// Exact current capability identity/type/revision; no blanket stale migration.
// AnyRevision: a restored document carries the ConfigRev of an earlier run, which
// says nothing about this one; the per-record identity, type and revision still do.
METHOD PRIVATE _M_ValidateSetShape : BOOL
VAR_INPUT
    Store : I_ConfigStore;
    Info : ST_ConfigSetInfo;
    AnyRevision : BOOL;
END_VAR
VAR
    expectedInfo : ST_ConfigSetInfo;
    expected : ST_ConfigRecord;
    record : ST_ConfigRecord;
    i : INT;
    j : INT;
    hits : INT;
END_VAR
_M_ValidateSetShape := FALSE;
IF (Store = 0) OR (Info.RootIdentity <> Status.Name)
OR (Info.SetSchema <> CONFIG_SET_SCHEMA)
OR (Info.RecordCount < 1) OR (Info.RecordCount > PL_Fraktal.MAX_SET_RECORDS) THEN
    _M_RejectConfigSet(Scope := Info.RootIdentity, Key := Info.SetName); RETURN;
END_IF
IF NOT AnyRevision AND ((Info.ConfigRev = 0) OR (Info.ConfigRev > ConfigRev)) THEN
    _M_RejectConfigSet(Scope := Info.RootIdentity, Key := Info.SetName); RETURN;
END_IF
IF NOT _snapshot.M_ReadInfo(SetName := '_validation', Info := expectedInfo) THEN RETURN; END_IF

FOR i := 1 TO Info.RecordCount DO
    IF NOT Store.M_ReadRecord(SetName := Info.SetName, Index := i, Record := record) THEN RETURN; END_IF
    hits := 0;
    FOR j := 1 TO expectedInfo.RecordCount DO
        _snapshot.M_ReadRecord(SetName := '_validation', Index := j, Record := expected);
        IF (record.Scope = expected.Scope) AND (record.WriteKey = expected.WriteKey) THEN
            IF (record.Kind <> expected.Kind) OR (record.ValueType <> expected.ValueType)
            OR (record.Revision <> expected.Revision) THEN
                _M_RejectConfigSet(Scope := record.Scope, Key := record.WriteKey); RETURN;
            END_IF
            hits := hits + 1;
        END_IF
    END_FOR
    IF hits <> 1 THEN
        _M_RejectConfigSet(Scope := record.Scope, Key := record.WriteKey); RETURN;
    END_IF
END_FOR
// Station sets may carry a subset; a Model bank or Line calendar is complete.
IF (Info.Kind <> E_ConfigKind.STATION_CFG) AND (Info.RecordCount <> expectedInfo.RecordCount) THEN
    _M_RejectConfigSet(Scope := Info.RootIdentity, Key := Info.SetName); RETURN;
END_IF
_M_ValidateSetShape := TRUE;
END_METHOD

// Append an inactive provider record. Live recipe and existing ordinals stay fixed.
METHOD CreateModel : BOOL
VAR_INPUT
    ModelCode : STRING(160);
    SourceIndex : UDINT;
    FromSet : BOOL;
    SetName : STRING(80);
END_VAR
VAR
    i : INT;
    info : ST_ConfigSetInfo;
    record : ST_ConfigRecord;
    source : I_ConfigStore;
    sourceName : STRING(80);
END_VAR
CreateModel := FALSE;
IF NOT _M_ConfigRestored() THEN
    RETURN;
END_IF
_exportNext := 0;
_M_SyncModelCatalog();
IF (_modelCatalog = 0) OR (_pModelRegion = 0) OR (_modelRegionSize < SIZEOF(UINT))
OR (ModelCode = '') OR (LEN(ModelCode) > 64) OR (AvailableModelCount >= ModelCapacity)
OR NOT Access.PermitsLogged(Gate := E_GatedAction.CONFIG_SET) THEN RETURN; END_IF
FOR i := 1 TO AvailableModelCount DO
    IF AvailableModels[i].ModelCode = ModelCode THEN RETURN; END_IF
END_FOR
// The exact bytes being validated are copied into the existing view buffer.
IF NOT _M_CaptureConfig(SetName := '_validation', Kind := E_ConfigKind.PAR_CFG,
        ModelIndex := SourceIndex) THEN RETURN; END_IF
source := _snapshot;
sourceName := '_validation';
IF FromSet THEN
    IF _configStore = 0 THEN RETURN; END_IF
    IF NOT _M_CopySet(SetName := SetName) THEN RETURN; END_IF
    IF NOT _loadSnapshot.M_ReadInfo(SetName := SetName, Info := info) THEN RETURN; END_IF
    IF info.Kind <> E_ConfigKind.PAR_CFG THEN RETURN; END_IF
    IF NOT _M_ValidateSetShape(Store := _loadSnapshot, Info := info,
            AnyRevision := FALSE) THEN RETURN; END_IF
    source := _loadSnapshot;
    sourceName := SetName;
END_IF
IF NOT source.M_ReadInfo(SetName := sourceName, Info := info) THEN RETURN; END_IF
MEMCPY(destAddr := ADR(_modelBuf), srcAddr := _pModelRegion, n := _modelRegionSize);
IF SourceIndex > 0 THEN
    IF AvailableModels[SourceIndex].ModelCode <> Model.ModelCode THEN
    IF NOT _modelProvider.Load(ModelCode := AvailableModels[SourceIndex].ModelCode,
            RecipeKey := _modelKey, pParCfg := ADR(_modelBuf), Size := _modelRegionSize) THEN RETURN; END_IF
    END_IF
END_IF
_pModelView := ADR(_modelBuf);
FOR i := 1 TO info.RecordCount DO
    IF NOT source.M_ReadRecord(SetName := sourceName, Index := i, Record := record) THEN EXIT; END_IF
    // A provider with one root record cannot clone another owner's recipe bank.
    IF NOT _M_OwnsModelRecord(Record := record) THEN EXIT; END_IF
    IF NOT Access.M_PermitsLevelLogged(Required := _M_DataLevelOf(TargetPath := record.Scope,
            WriteKey := record.WriteKey, ForWrite := FALSE)) THEN EXIT; END_IF
    IF NOT Access.M_PermitsLevelLogged(Required := _M_DataLevelOf(TargetPath := record.Scope,
            WriteKey := record.WriteKey, ForWrite := TRUE)) THEN EXIT; END_IF
    IF NOT SUPER^.M_ApplyConfigWrite(Scope := record.Scope, WriteKey := record.WriteKey,
            Revision := record.Revision, TextValue := record.ValueText, RootReady := TRUE) THEN EXIT; END_IF
END_FOR
_pModelView := 0;
IF i <= info.RecordCount THEN RETURN; END_IF
CreateModel := _modelCatalog.M_CreateModel(ModelCode := ModelCode, RecipeKey := _modelKey,
    pData := ADR(_modelBuf), Size := _modelRegionSize);
IF CreateModel THEN
    _M_SyncModelCatalog();
    _M_MarkPersistPending();
END_IF
END_METHOD

METHOD ExportCurrentConfig : BOOL
VAR_INPUT
    SetName : STRING(80);
    Kind : E_ConfigKind;
    ModelIndex : UDINT;
    Token : STRING(160);
END_VAR
VAR
    info : ST_ConfigSetInfo;
    record : ST_ConfigRecord;
    i : INT;
END_VAR
ExportCurrentConfig := FALSE;
_exportNext := 0;
ConfigSetDocument := '';
ConfigSetDocumentLines := 0;
IF (Token = '') OR Access.ReqLogout
OR NOT Access.Permits(Gate := E_GatedAction.CONFIG_SET) THEN RETURN; END_IF
IF NOT _M_CaptureConfig(SetName := SetName, Kind := Kind, ModelIndex := ModelIndex) THEN RETURN; END_IF
_snapshot.M_ReadInfo(SetName := SetName, Info := info);
FOR i := 1 TO info.RecordCount DO
    _snapshot.M_ReadRecord(SetName := SetName, Index := i, Record := record);
    IF NOT Access.M_PermitsLevel(Required := _M_DataLevelOf(TargetPath := record.Scope,
            WriteKey := record.WriteKey, ForWrite := FALSE)) THEN RETURN; END_IF
END_FOR
_exportToken := Token;
_exportSession := Access.SessionGeneration;
_exportName := SetName;
_exportNext := 1;
ConfigSetDocument := _setJson.M_Header(Info := info);
ConfigSetDocumentLine := 0;
ConfigSetDocumentLines := info.RecordCount;
ExportCurrentConfig := ConfigSetDocument <> '';
END_METHOD

METHOD PRIVATE _M_ExportSnapshotLine : BOOL
VAR_INPUT
    SetName : STRING(80);
    Line : INT;
    Token : STRING(160);
END_VAR
VAR
    info : ST_ConfigSetInfo;
    record : ST_ConfigRecord;
END_VAR
_M_ExportSnapshotLine := FALSE;
ConfigSetDocument := '';
ConfigSetDocumentLines := 0;
IF (_exportNext = 0) OR (Line <> _exportNext) OR (Token <> _exportToken)
OR (_exportSession <> Access.SessionGeneration) OR (SetName <> _exportName)
OR Access.ReqLogout
OR NOT Access.Permits(Gate := E_GatedAction.CONFIG_SET) THEN
    _exportNext := 0; RETURN;
END_IF
IF NOT _snapshot.M_ReadInfo(SetName := SetName, Info := info)
OR NOT _snapshot.M_ReadRecord(SetName := SetName, Index := Line, Record := record) THEN
    _exportNext := 0; RETURN;
END_IF
IF NOT Access.M_PermitsLevel(Required := _M_DataLevelOf(TargetPath := record.Scope,
        WriteKey := record.WriteKey, ForWrite := FALSE)) THEN
    _exportNext := 0; RETURN;
END_IF
ConfigSetDocument := _setJson.M_Record(Record := record);
ConfigSetDocumentLine := Line;
ConfigSetDocumentLines := info.RecordCount;
_exportNext := _exportNext + 1;
IF Line = info.RecordCount THEN _exportNext := 0; END_IF
_M_ExportSnapshotLine := ConfigSetDocument <> '';
END_METHOD

END_FUNCTION_BLOCK

(* stored: Version 1.1.0.1, ProductVersion 3.1.4024.16
   POU FB_UnitBase: Id {116d9026-fbad-4cf8-8b52-50d17613c706}, SpecialFunc None
   Method _M_AddReason: Id {63c5e93f-708a-4c3a-aa1b-ee43d815fb4a}
   Method _M_AppendInterlocks: Id {2bc971ff-4cee-49e6-a29f-4f727818205b}
   Method _M_AppendManualInterlocks: Id {c18caeb9-871a-4a4c-aad2-2711e3ced37a}
   Method _M_AppendDecisionInterlocks: Id {bbac41d9-35ba-4800-af52-51cd30b49db7}
   Method _M_AskDecision: Id {4e23ce8a-174c-4663-9cbe-be702ba37032}
   Method _M_ClearDecisionState: Id {db09e3d9-4427-4607-8a90-66b39812e37b}
   Method _M_DecisionCyclic: Id {ff058255-d664-4ce3-986d-8ad7a970388c}
   Method _M_DecisionMatches: Id {2ca48458-620f-4a17-b6d1-b5680778bd4e}
   Method _M_LogDecision: Id {eb357477-2029-4b6d-8688-04dc5df5e04b}
   Method _M_ValidateDecision: Id {1229fbc9-7dc8-4907-b878-f6af733f2c09}
   Method _M_Await: Id {098638cb-fc78-4032-9954-0ceffe6b565c}
   Method _M_CascadeMode: Id {3ac20481-72c5-4cd1-88e5-b9f7eb433162}
   Method _M_ClearPending: Id {cb01b1f4-f591-43f7-a826-970be7300b04}
   Method _M_AuditHmiAccepted: Id {f8865f87-3ae7-472e-b775-3408513a4586}
   Method _M_OwnsModulePath: Id {9b8c6045-f404-4484-937e-b0a8f749d8fd}
   Method _M_EndOfCycle: Id {9824e487-d8d3-4cb9-8c78-a6d2fc09a62d}
   Method _M_HandleHmiRequest: Id {63ae9d50-339f-4904-a8ec-81f853aed962}
   Method _M_HostEvent: Id {76fb49ac-f9ea-4e53-8db6-e7e4e756fd84}
   Method _M_InitModePolicy: Id {df8ba8da-c8fa-411c-85c1-392b353d5cfd}
   Method _M_OeeCompute: Id {2991f1a8-70f1-48a9-aa83-352243818d0a}
   Method _M_OeeUpdate: Id {8a4f011d-5d7a-4935-ad26-8a5fbcf63643}
   Method _M_PartAborted: Id {a55c31e8-06f9-4d10-8c26-4e83b7d5c1f2}
   Method _M_PartEvent: Id {f18c2d47-9b53-4e6a-8c02-3a71d5f0b429}
   Method _M_PartProcessed: Id {e91b5a02-73df-4f16-a8d4-1c30fe8a97d2}
   Method _M_PartReceived: Id {58c0a7d9-14be-4f22-8d6a-9b2ef4c1e370}
   Method _M_PartRecord: Id {7be4f6a3-1d20-4c8e-be55-f2a09318d67c}
   Method _M_PartStarted: Id {02a97d1c-6bb5-4f80-9d34-c58b12f04ae6}
   Method _M_PublishStatus: Id {02d44270-09e8-4bc1-97fd-f43dd3fc44f2}
   Method _M_PushHistory: Id {3f9af757-7ef5-4499-8b8d-04dcd97acc93}
   Method _M_RaiseMaintenance: Id {c92e4b71-6d05-4f88-9e3a-2b17d4c8a054}
   Method _M_RouteConfigWrite: Id {4e524daf-e482-4764-8639-e58c1f363aa3}
   Method _M_WriteBaseConfig: Id {c30f39b4-eae4-421d-a415-c6dc3b402679}
   Method _M_RouteForceChannel: Id {301182d5-8822-451a-950c-49d23daf4640}
   Method _M_RouteManual: Id {9fa4e2c2-3f5f-4681-aed5-559f1df0d2c6}
   Method _M_RecordSequenceStep: Id {bae7334e-b67d-46db-a917-aa05f1522e0f}
   Method _M_ResetSequenceRows: Id {3a7e979a-9c02-4e58-aa36-f0627902f8fb}
   Method _M_SequenceAnnotate: Id {981fa92c-f12b-4972-9483-880edfae72c8}
   Method _M_SequenceAnnotationClear: Id {7256d50d-cf16-4906-8e35-fd394563602f}
   Method _M_SetStep: Id {1066dd3c-baf2-43ea-91d5-309ad4ca7878}
   Method _M_StallWalk: Id {ee453cd4-7027-4207-b43e-f1a12367922c}
   Method _M_StepGate: Id {853d1e75-22c1-46fb-9a92-007882839a98}
   Method _M_Supports: Id {5285aa9e-3e18-4090-bed9-0119293228bb}
   Method _M_SupportsRunStyle: Id {f4e81ed4-d8b0-494c-bd7a-6b417d6219cf}
   Method _M_TakeDecision: Id {e2e1443d-0421-4608-8ae5-b7bb44177b3c}
   Method CountGood: Id {852e951b-039f-45bd-80a3-6417310e2406}
   Method CountNok: Id {a686f5b6-4c90-4e12-9d98-fa111d14dfe8}
   Method CountRework: Id {5c8e02d7-9a41-4f36-8b52-e04a71c6d983}
   Method M_AppendConfig: Id {29c7f5d4-0b81-4ae3-9762-84f6d013ba58}
   Method SetConfigStore: Id {1f6b90d4-38a2-4c57-9e01-b47d2c85a3f6}
   Method SetPersistMedium: Id {90949ce0-2dde-4312-82c9-779c3854619d}
   Method SetConfigPersistence: Id {a5c37e08-9412-4bd6-83f9-6e05b17c94a2}
   Method SetConfigPersistWindow: Id {5db2740a-9e18-4c63-b0f5-8a2914e7c036}
   Method SetConfigRestorePolicy: Id {72e4a1b9-c530-46df-8127-93b605ea4d78}
   Method _M_MarkPersistPending: Id {6d09fb35-2a84-41ce-b7f0-58d2e1937a4b}
   Method _M_ConfigPersistFailed: Id {3a81c6e7-40b2-4d95-916f-c82705bd4e13}
   Method _M_ConfigPersistCyclic: Id {9c0d4318-b7a5-42e6-8f13-05ea7c9b2d40}
   Method _M_ConfigRestored: Id {c723ef57-9111-489a-87e1-2e9e98d880fe}
   Method _M_LiveCyclic: Id {aad84a07-4f6e-415a-a949-44d11c57baf2}
   Method _M_LiveReadFailed: Id {c1b391b8-49e2-405b-9490-706629300cca}
   Method _M_LivePassFailed: Id {3fff4db1-40c0-4916-a009-f750b7b16137}
   Method _M_LiveItemUsed: Id {2d7178d4-917d-4032-9b90-b6d8a8215873}
   Method _M_LiveKey: Id {77a63a7d-cd03-4447-be78-e758d5ef1591}
   Method _M_LiveModelsKept: Id {166da471-060a-4724-bca3-30a7b039d62b}
   Method _M_LiveRestoreItem: Id {b20141f1-cfd8-47d0-b996-33c491a3a370}
   Method _M_LiveApply: Id {031ae06a-8d84-4843-bce8-ed6d53fdc0d1}
   Method _M_ModelIndexOf: Id {055b30d9-edd2-408c-ae7f-7015e649658e}
   Method _M_DrainRestoreLoss: Id {0b7e5294-16ad-43c1-a8f6-249d038be715}
   Method _M_AnnounceRestoreLoss: Id {77125c95-ab46-4aaa-9f22-3a07f8e7fd8f}
   Method AcknowledgeConfigRestore: Id {e18c47b3-5029-4ed6-9a71-b3406fc25d89}
   Method _M_RejectConfigSet: Id {5f2a90c6-8b41-4d73-bec0-172e845f39ab}
   Method _M_SetOpAllowed: Id {3d70b95e-c284-41f0-86ba-9e15c703da42}
   Method DeleteConfigSet: Id {e533f05f-2594-42e8-8c99-81d549fc4090}
   Method _M_DataLevelOf: Id {181e4912-d325-4208-982a-bde235412443}
   Method M_DeclareDataClass: Id {b9a4a5ae-9fab-42bd-bc82-7e32dffbd2a9}
   Method SetDataClassLevel: Id {047e7f36-274a-4350-8ad6-b77d4f72cc43}
   Method _M_IsLineKey: Id {59358b2d-9028-416d-b8b1-1699a6cd425f}
   Method M_ApplyConfigWrite: Id {09d95f4a-6281-4745-bbd6-78a379c3dcc0}
   Method M_StageConfigWrite: Id {c033d610-c896-4206-a3ad-81018a4dd465}
   Method M_ApplyCapture: Id {e2ff8450-6122-448e-b867-574b3000edfa}
   Method M_ConfigAccessOf: Id {b5882f05-b837-4f44-ba08-a65bdacad4e2}
   Method M_RegisterModelData: Id {9e19e4d6-5131-4b98-84c6-f84c0e107ced}
   Method _M_OpenModelView: Id {93ccf92c-d752-48c8-af0b-7941488b3430}
   Method WriteModelConfig: Id {2a0d9e3e-ba70-4e09-955f-cec98e39642e}
   Method M_AppendModelConfig: Id {0e6d90bf-ad76-4384-ab12-1767af3d1a4f}
   Method _M_SaveModelData: Id {614f64a8-a7bb-415b-89b6-cd5638516728}
   Method SetLine: Id {b3e3c826-6085-43fe-ab9e-5ee8d63ca7f0}
   Method M_ShiftTick: Id {4606cb81-948b-4fb3-a998-828e0341cdfd}
   Method _M_CloseShift: Id {3589014a-a797-47c8-9c22-164193338f8a}
   Method SaveConfigSet: Id {8a4d1e07-63b9-4c25-90fd-e7285a1cb046}
   Method LoadConfigSet: Id {c93f5b28-047e-41da-b6c1-5820ae74f3d9}
   Method _M_ApplySet: Id {f003cd3e-e4eb-4ec5-b15b-c46e595f4b79}
   Method _M_StageOneRecord: Id {b6014e8d-72c3-49a5-80fe-c1738d92406b}
   Method _M_ConfigSetHalfApplied: Id {47db6015-9a2e-4c38-b7f0-d5216e409a83}
   Method ListConfigSets: Id {2e85d740-c6b1-4930-a5df-08417b3ce629}
   Method ExportConfigSetLine: Id {6c1908fe-b432-4a07-95d8-e2603ba7145c}
   Method ImportConfigSetLine: Id {d0a76321-8e54-4bc9-97a2-3f16054eb7d8}
   Method ImportConfigSetPiece: Id {fe4a451b-e9cc-440c-9ade-c56031168c94}
   Method M_SequenceAskDecision: Id {099b4f9d-bc09-44d1-a376-b2e504dbb242}
   Method M_SequenceAwait: Id {c61669f7-ff2f-475c-915e-c23e673ae50d}
   Method M_SequenceClearDecision: Id {f5e88d63-dd7e-45c7-8fcc-149437ebcb66}
   Method M_SequenceComplete: Id {94f85c2c-bf7e-4679-9ad7-df299f9443e9}
   Method M_SequenceCountGood: Id {7ac5d064-bbc3-4e23-a999-5b1106c18501}
   Method M_SequenceEndOfCycle: Id {2465831e-ce6a-49ba-894a-d94a6e5b730d}
   Method M_SequenceFault: Id {6dcf30ea-273a-4919-b53c-93ee346a0722}
   Method M_SequencePartProcessed: Id {f3fe635f-f0ef-4b80-918f-2af11c08a018}
   Method M_SequencePartReceived: Id {9576ad5e-fef2-4d71-bd9f-075e2fbf7f48}
   Method M_SequencePartRecord: Id {272bc8d6-51f1-4e02-a0f6-834fc34cf443}
   Method M_SequencePartStarted: Id {c34399dc-9677-414b-87a7-da41fec81ce1}
   Method M_SequenceRegister: Id {9c12e1e0-2b54-4710-a719-b7dbb939da2c}
   Method _M_BeginSequenceScan: Id {90d173ad-1ac7-44ea-8963-773d827fd02e}
   Method _M_RestartSequences: Id {a7179c76-6bab-4060-a5d3-1d37fa9ff028}
   Method OnAbort: Id {045fbfe7-105f-49b4-bf25-f60661612052}
   Method OnAbortInError: Id {f7465218-0d83-46fd-a26a-73b938ae69a7}
   Method M_SequenceWarn: Id {75ce463f-f749-4a05-8c5e-fea3607d380d}
   Method M_SequenceRaise: Id {0bee2dd9-d8a8-4946-b400-dc31452b748f}
   Method _M_ResumeSequencesAfterError: Id {f331535e-fb67-4439-a403-97a206176d31}
   Method M_SequenceSetStep: Id {cd33b52b-b93d-4827-921b-0507be840f66}
   Method M_SequenceStepGate: Id {4300b99e-dada-4558-9a7d-f357bb3b59db}
   Method M_SequenceStopNow: Id {5e2a91d7-38c4-4b0f-a6e8-74d19c2b50f3}
   Method M_SequenceStopPending: Id {9b04e7c1-52d8-4f36-8a92-1c65fd83a247}
   Method M_SequenceTakeDecision: Id {a0cad3a5-90f7-4b63-9dfc-d75845d8e702}
   Method ManualHeldTo: Id {9a41c8e0-5b73-4d26-81fa-06e5327d94b1}
   Method _M_RouteHeld: Id {3c78e05b-1246-4a9d-b0e7-52f8146c93da}
   Method _M_ChartRevCyclic: Id {b40f7e26-95a1-4d83-b217-0c6e59a71e34}
   Method _M_HeldCyclic: Id {d51937ae-64c2-408f-9b13-27e0a4586cf7}
   Method ManualCommandTo: Id {4de99325-2725-4710-8292-b2f11cd5c61c}
   Property ModeActive: Id {cadd011f-36e9-480f-9687-f764db6a93a1}
   Get Get: Id {480f723e-9802-4414-9cf5-b9bf28538b7e}
   Property ModelCode: Id {52be901d-358c-42d1-8de9-24cabf037285}
   Get Get: Id {d1228112-dc00-4a78-8d96-06a0aa3db5e2}
   Property ModuleType: Id {19c4f994-fbe0-4e50-80d5-d89b1a1fb1fa}
   Get Get: Id {e694d09e-29b1-48cc-b1e6-0d26ae208150}
   Method OnCyclic: Id {833bee58-3464-412f-8fa3-37fa398fef55}
   Method _M_HighestSeverity: Id {06beeb70-94f2-4095-9daa-a1af1fd36a20}
   Method RequestLampTest: Id {0a1df30a-092c-4f3f-91a5-1af799e7cb11}
   Method SetSignalTowerConfig: Id {93bf4461-f32d-446c-ac46-8d0b800f56d9}
   Method SetSystemHealth: Id {f544458e-b3ee-4aad-ac8d-2565c5120fa3}
   Method OnInit: Id {c11afaa2-3957-4d40-8695-293ff272dfc1}
   Method OnModeChanged: Id {4307796c-f352-4515-b104-1671ef41b10c}
   Method OnCommandStart: Id {4698d7ce-6d4c-492c-9ead-e072c285ae34}
   Method OnModeExit: Id {d824838b-6d6c-4575-ade3-00f3815d6c9e}
   Method OperatorReset: Id {86e0365e-0665-41e9-b6f4-1156fe1cf971}
   Method _M_RecoverState: Id {2d0b998f-abd6-473c-8cb5-b6b35c39d09a}
   Method OnOperatorReset: Id {ad173c6c-fa19-47ee-a347-f5b5e0c7654a}
   Method RequestLocalReset: Id {2ac5c84b-a29d-437a-b5c9-0d4b5d278812}
   Method RegisterAvailableModel: Id {651bb1e1-71c6-4fb4-a063-4ea057e752cf}
   Method RequestControlPower: Id {cb696b98-d3f2-48ed-8f23-09e45169ea5f}
   Method SubmitDecision: Id {70347f2b-2424-4514-beb7-8788c8d00fca}
   Method SetAccessLevel: Id {a2b5995c-ea0a-4911-83f3-0a5e24269563}
   Method SetSessionTimeout: Id {e8244b36-18c3-4b2a-8ef7-db39a1dfa257}
   Method WriteConfig: Id {3e40e571-e45f-4204-a5d3-c9907077e8b2}
   Method CaptureConfig: Id {6657c29b-54a9-410f-b368-d4a1ad1bb646}
   Method SetEngineeringMode: Id {28e702f3-e7d8-4e5a-8206-7208a16b6696}
   Method M_ForcePermitted: Id {b9d8bf79-0c6d-4741-99f8-f427bda243e9}
   Method _M_EngineeringCyclic: Id {0b6876ea-bb0c-4e77-ab09-61eab13a8627}
   Method ForceChannel: Id {8bf9fd9d-8084-4dbf-b41b-c60e5e0cc995}
   Method ReleaseReportAction: Id {b52c134c-be50-4c5c-b4df-ad025ff72931}
   Method ReleaseReportManual: Id {9e9f491d-e5a8-435c-bc95-8f93e8c3530b}
   Method ReleaseReportStart: Id {c78c7568-83f2-4d9d-9ae3-f47850cbc022}
   Method ResetOee: Id {76d2024b-e4e9-424e-bbf4-fcfd488c8439}
   Method SetHoldRun: Id {fbc37d38-8939-4f18-83b4-eb1341e2b47b}
   Method SetIdealCycle: Id {21a43259-c0d5-420f-993f-704ffad3d187}
   Method SetMode: Id {7da8ba28-e926-421f-9272-a6c57a552866}
   Method SetModel: Id {6a7ae71f-5111-44b3-bfc5-fd8bfdcd3719}
   Method M_PublishMaterialChanged: Id {27225091-fd15-48c0-a242-131de64ab93c}
   Method M_PublishToolChanged: Id {cc18bd59-d3df-4af3-a8b4-e56788466431}
   Method M_SetHostEventSink: Id {c075ef1c-ce1a-4aec-9cd4-f8cc578ba7b2}
   Method SetPartCarrier: Id {6a3e9c15-2f84-4b0d-9c17-d84f5e21ab63}
   Method SetRunStyle: Id {f598b9ad-9cb8-47de-920d-91798ab2094a}
   Method ShelveAlarm: Id {254b8716-80f2-462f-8e49-d89ea86b5224}
   Method Start: Id {cf23e563-6a38-441b-bf71-cf054a5930b3}
   Method StepRequest: Id {64e64e1a-0c5a-460b-882a-ab14da4420e6}
   Method Stop: Id {a7c9b0f8-857c-458d-afc6-9746ac288208}
   Property StopPending: Id {f114fa1a-de45-4aa0-be5b-cf63c773b8b7}
   Get Get: Id {135b3f46-0e90-48aa-8ac1-6493d51adeb3}
   Method UnshelveAlarm: Id {f39e65ca-0fee-42d8-be9a-7e2098b02e14}
   Method _M_SyncModelCatalog: Id {b4da8c6b-131b-4566-b7f8-2b4dad9efb38}
   Method _M_OwnsModelRecord: Id {49fcf615-a1bb-43fd-a838-ed96547c3417}
   Method _M_CopySet: Id {c431d797-d523-47f2-b0d9-d224d1cd55f1}
   Method _M_CaptureConfig: Id {3631f460-c887-48c6-a7aa-a345c944f785}
   Method _M_CaptureInto: Id {29414adf-e5e0-41d7-bc26-9a37ff215723}
   Method _M_ValidateSetShape: Id {6aad96f0-b145-4801-97ec-47145f5fcee6}
   Method CreateModel: Id {cc3c11aa-cac7-4411-9bca-a1f3f1acdb30}
   Method ExportCurrentConfig: Id {6b0ac5cd-01e5-48b3-8c05-7e155068df6f}
   Method _M_ExportSnapshotLine: Id {7d34463f-e19c-4d8f-bed9-72b0b2732824} *)
